Fanuc KAREL source: KA00072.KL

PROGRAM KA00072
%NOLOCKGROUP
VAR
  SRC: XYZWPR
  DST: ARRAY[2] OF SHORT
BEGIN
  SRC.X = 1.0
  DST[1] = SRC
END KA00072
